DATA_BLOCK "Current_state_of_Bay1"
{ S7_Optimized_Access := 'TRUE' }
VERSION : 0.1
NON_RETAIN
   VAR
      Bay1 : Array[0..3, 0..11] of UInt;
   END_VAR


BEGIN
   Bay1[0,0] := 555;
   Bay1[0,1] := 556;
   Bay1[0,2] := 0;
   Bay1[0,3] := 0;
   Bay1[0,4] := 0;
   Bay1[0,5] := 0;
   Bay1[0,6] := 0;
   Bay1[0,7] := 0;
   Bay1[0,8] := 0;
   Bay1[0,9] := 0;
   Bay1[0,10] := 0;
   Bay1[0,11] := 0;
   Bay1[1,0] := 557;
   Bay1[1,1] := 0;
   Bay1[1,2] := 0;
   Bay1[1,3] := 0;
   Bay1[1,4] := 0;
   Bay1[1,5] := 0;
   Bay1[1,6] := 0;
   Bay1[1,7] := 0;
   Bay1[1,8] := 0;
   Bay1[1,9] := 0;
   Bay1[1,10] := 0;
   Bay1[1,11] := 0;
   Bay1[2,0] := 0;
   Bay1[2,1] := 0;
   Bay1[2,2] := 0;
   Bay1[2,3] := 0;
   Bay1[2,4] := 0;
   Bay1[2,5] := 0;
   Bay1[2,6] := 0;
   Bay1[2,7] := 0;
   Bay1[2,8] := 0;
   Bay1[2,9] := 0;
   Bay1[2,10] := 0;
   Bay1[2,11] := 0;
   Bay1[3,0] := 0;
   Bay1[3,1] := 0;
   Bay1[3,2] := 0;
   Bay1[3,3] := 0;
   Bay1[3,4] := 0;
   Bay1[3,5] := 0;
   Bay1[3,6] := 0;
   Bay1[3,7] := 0;
   Bay1[3,8] := 0;
   Bay1[3,9] := 0;
   Bay1[3,10] := 0;
   Bay1[3,11] := 0;

END_DATA_BLOCK

